// TIA Portal V21 export
// export: Created 2026-11-21T13:24:04.6188738Z, ExportSetting WithDefaults, DisplayName Totally Integrated Automation Portal, DisplayVersion V21, DisplayName STEP 7 Professional, DisplayVersion V21, DisplayName STEP 7 Safety, DisplayVersion V21, DisplayName Tech WebApplication, DisplayVersion V21, DisplayName WinCC Basic/Comfort/Advanced, DisplayVersion V21, DisplayName WinCC Unified, DisplayVersion V21
FUNCTION_BLOCK "Guard"   // FB5, F_FBD
{ S7_Optimized_Access := 'TRUE' }
VERSION : 0.1
// A guard door: open while its switch is not closed.
// stored: AutoNumber true, IsIECCheckEnabled false, UDAEnableTagReadback false
   VAR_INPUT
      closed : Bool;
   END_VAR
   VAR_OUTPUT
      open : Bool;
   END_VAR
BEGIN

REGION Network 1: Open guard
   // The guard is open while its switch is not closed.
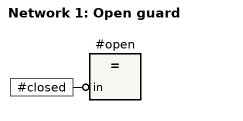
   #open := NOT #closed;
END_REGION
END_FUNCTION_BLOCK
